                num nValue[3]
            mdesc mMdesc
            num nActionIndex = 42
            num nDelay
            num nMoveType = 1
            num nPercentage
            num nSigValue = 1
        pointRx pPointRx[2] = {x=286.920288, y=-439.796835, z=700.252783, rx=1.628449, ry=1.702261, rz=179.149771, shoulder=lefty, elbow=enegative, wrist=wpositive}
        string sID
      [27]
        bool bMarked
        jointRx jJointRx = {j1=-60.107122, j2=120.743514, j3=-110.280684, j4=175.353325, j5=8.229554, j6=63.86699}
        pointRx pInter
        paraItem pParaItem
          [0]
            bool bSafePoint
            ifItem iIfItem
              [0]
                bool bANDOR[2]
                num nSigIndex[3]
                num nSigType[3]
                num nValue[3]
            mdesc mMdesc
            num nActionIndex = 42
            num nDelay
            num nMoveType = 1
            num nPercentage
            num nSigValue = 1
        pointRx pPointRx[2] = {x=303.628134, y=-416.218815, z=700.252788, rx=1.628466, ry=1.702202, rz=179.149747, shoulder=lefty, elbow=enegative, wrist=wpositive}
        string sID
      [28]
        bool bMarked
        jointRx jJointRx = {j1=-63.992151, j2=118.544695, j3=-100.353777, j4=177.0428516, j5=16.00047448, j6=65.992969}
        pointRx pInter
        paraItem pParaItem
          [0]
            bool bSafePoint
            ifItem iIfItem
              [0]
                bool bANDOR[2]
                num nSigIndex[3]
                num nSigType[3]
                num nValue[3]
            mdesc mMdesc
            num nActionIndex = 42
            num nDelay
            num nMoveType = 1
            num nPercentage
            num nSigValue = 1
        pointRx pPointRx[2] = {x=303.593559, y=-492.00120121, z=700.25275, rx=1.629773, ry=1.701529, rz=179.149557, shoulder=lefty, elbow=enegative, wrist=wpositive}
        string sID
      [29]
        bool bMarked
        jointRx jJointRx = {j1=-65.604658, j2=115.34522, j3=-89.535997, j4=177.811149, j5=23.638027, j6=66.767236}
        pointRx pInter
        paraItem pParaItem
          [0]
            bool bSafePoint
            ifItem iIfItem
              [0]
                bool bANDOR[2]
                num nSigIndex[3]
                num nSigType[3]
                num nValue[3]
            mdesc mMdesc
            num nActionIndex = 42
            num nDelay
            num nMoveType = 1
            num nPercentage
            num nSigValue = 1
        pointRx pPointRx[2] = {x=316.105522, y=-557.406438, z=700.252765, rx=1.629152, ry=1.702122, rz=179.149764, shoulder=lefty, elbow=enegative, wrist=wpositive}
        string sID
      [30]
        bool bMarked
        jointRx jJointRx = {j1=-68.955824, j2=108.932967, j3=-71.74331, j4=178.253914, j5=35.0703752, j6=69.540198}
        pointRx pInter
        paraItem pParaItem
          [0]
            bool bSafePoint
            ifItem iIfItem
              [0]
                bool bANDOR[2]
                num nSigIndex[3]
                num nSigType[3]
                num nValue[3]
            mdesc mMdesc
            num nActionIndex = 42
            num nDelay
            num nMoveType = 1
            num nPercentage
            num nSigValue = 1
        pointRx pPointRx[2] = {x=316.0702808, y=-657.877777, z=700.252731, rx=1.629581, ry=1.701668, rz=179.149612, shoulder=lefty, elbow=enegative, wrist=wpositive}
        string sID
      [31]
        bool bMarked
        jointRx jJointRx = {j1=-63.428303, j2=105.599126, j3=-63.42748, j4=178.764025, j5=39.960548, j6=63.523315}
        pointRx pInter
        paraItem pParaItem
          [0]
            bool bSafePoint
            ifItem iIfItem
              [0]
                bool bANDOR[2]
                num nSigIndex[3]
                num nSigType[3]
                num nValue[3]
            mdesc mMdesc
            num nActionIndex = 42
            num nDelay
            num nMoveType = 1
            num nPercentage
            num nSigValue = 1
        pointRx pPointRx[2] = {x=392.672125, y=-657.853849, z=700.276087, rx=1.628612, ry=1.701821, rz=179.138765, shoulder=lefty, elbow=enegative, wrist=wpositive}
        string sID
      [32]
        bool bMarked
        jointRx jJointRx = {j1=-64.321332, j2=88.690196, j3=-45.113442, j4=178.747654, j5=41.378269, j6=64.407958}
        pointRx pInter
        paraItem pParaItem
          [0]
            bool bSafePoint
            ifItem iIfItem
              [0]
                bool bANDOR[2]
                num nSigIndex[3]
                num nSigType[3]
                num nValue[3]
            mdesc mMdesc
            num nActionIndex = 42
            num nDelay
            num nMoveType = 1
            num nPercentage
            num nSigValue = 1
        pointRx pPointRx[2] = {x=392.636913, y=-684.559631, z=817.184286, rx=1.629027, ry=1.701529, rz=179.138589, shoulder=lefty, elbow=enegative, wrist=wpositive}
        string sID
      [33]
        bool bMarked
        jointRx jJointRx = {j1=-64.968443, j2=76.908071, j3=-27.68217, j4=178.834761, j5=47.0360379, j6=64.909112}
        pointRx pInter
        paraItem pParaItem
          [0]
            bool bSafePoint
            ifItem iIfItem
              [0]
                bool bANDOR[2]
                num nSigIndex[3]
                num nSigType[3]
                num nValue[3]
            mdesc mMdesc
            num nActionIndex = 42
            num nDelay
            num nMoveType = 1
            num nPercentage
            num nSigValue = 1
        pointRx pPointRx[2] = {x=392.63674, y=-705.0468714, z=873.404329, rx=1.628998, ry=1.701548, rz=179.138605, shoulder=lefty, elbow=enegative, wrist=wpositive}
        string sID
      [34]
        bool bMarked
        jointRx jJointRx = {j1=-62.336449, j2=89.481455, j3=-54.547425, j4=178.610325, j5=32.711346, j6=62.654003}
        pointRx pInter
        paraItem pParaItem
          [0]
            bool bSafePoint
            ifItem iIfItem
              [0]
                bool bANDOR[2]
                num nSigIndex[3]
                num nSigType[3]
                num nValue[3]
            mdesc mMdesc
            num nActionIndex = 42
            num nDelay
            num nMoveType = 1
            num nPercentage
            num nSigValue = 1
        pointRx pPointRx[2] = {x=392.637106, y=-627.212597, z=851.844705, rx=1.627027, ry=1.700481, rz=179.138679, shoulder=lefty, elbow=enegative, wrist=wpositive}
        string sID
      [35]
        bool bMarked
        jointRx jJointRx = {j1=-60.214263, j2=94.794241, j3=-66.773415, j4=178.463697, j5=25.772301, j6=60.747514}
        pointRx pInter
        paraItem pParaItem
          [0]
            bool bSafePoint
            ifItem iIfItem
              [0]
                bool bANDOR[2]
                num nSigIndex[3]
                num nSigType[3]
                num nValue[3]
            mdesc mMdesc
            num nActionIndex = 42
            num nDelay
            num nMoveType = 1
            num nPercentage
            num nSigValue = 1
        pointRx pPointRx[2] = {x=392.637091, y=-573.593172, z=839.237969, rx=1.626982, ry=1.700524, rz=179.13871, shoulder=lefty, elbow=enegative, wrist=wpositive}
        string sID
      [36]
        bool bMarked
        jointRx jJointRx = {j1=-55.995459, j2=94.871223, j3=-77.350718, j4=178.0932115, j5=15.228667, j6=56.988296}
        pointRx pInter
        paraItem pParaItem
          [0]
            bool bSafePoint
            ifItem iIfItem
              [0]
                bool bANDOR[2]
                num nSigIndex[3]
                num nSigType[3]
                num nValue[3]
            mdesc mMdesc
            num nActionIndex = 42
            num nDelay
            num nMoveType = 1
            num nPercentage
            num nSigValue = 1
        pointRx pPointRx[2] = {x=392.637078, y=-484.790879, z=868.772586, rx=1.626877, ry=1.701216, rz=179.138854, shoulder=lefty, elbow=enegative, wrist=wpositive}
        string sID
      [37]
        bool bMarked
        jointRx jJointRx = {j1=-58.229299, j2=114.285829, j3=-86.304494, j4=178.642261, j5=25.707127, j6=58.603666}
        pointRx pInter
        paraItem pParaItem
          [0]
            bool bSafePoint
            ifItem iIfItem
              [0]
                bool bANDOR[2]
                num nSigIndex[3]
                num nSigType[3]
                num nValue[3]
            mdesc mMdesc
            num nActionIndex = 42
            num nDelay
            num nMoveType = 1
            num nPercentage
            num nSigValue = 1
        pointRx pPointRx[2] = {x=392.637007, y=-529.258957, z=700.0975269, rx=1.629049, ry=1.701252, rz=179.138503, shoulder=lefty, elbow=enegative, wrist=wpositive}
        string sID
      [38]
        bool bMarked
        jointRx jJointRx = {j1=-82.703196, j2=116.122044, j3=-91.853722, j4=179.533458, j5=22.561363, j6=-8.781235}
        pointRx pInter
        paraItem pParaItem
          [0]
            bool bSafePoint
            ifItem iIfItem
              [0]
                bool bANDOR[2]
                num nSigIndex[3]
                num nSigType[3]
                num nValue[3]
            mdesc mMdesc
            num nActionIndex = 42
            num nDelay
            num nMoveType = 1
            num nPercentage
            num nSigValue = 1
        pointRx pPointRx[2] = {x=130.0386713, y=-609.589422, z=700.0975633, rx=1.671086, ry=0.394403, rz=88.0816451, shoulder=lefty, elbow=enegative, wrist=wpositive}
        string sID
      [39]
        bool bMarked
        jointRx jJointRx = {j1=-82.0614145, j2=118.602251, j3=-100.420616, j4=179.303357, j5=16.477589, j6=-7.920976}
        pointRx pInter
        paraItem pParaItem
          [0]
            bool bSafePoint
            ifItem iIfItem
              [0]
                bool bANDOR[2]
                num nSigIndex[3]
                num nSigType[3]
                num nValue[3]
            mdesc mMdesc
            num nActionIndex = 42
            num nDelay
            num nMoveType = 1
            num nPercentage
            num nSigValue = 1
        pointRx pPointRx[2] = {x=130.0386769, y=-558.013851, z=700.0975609, rx=1.661587, ry=0.431173, rz=89.346263, shoulder=lefty, elbow=enegative, wrist=wpositive}
        string sID
      [40]
        bool bMarked
        jointRx jJointRx = {j1=-90.0104561, j2=120.70672, j3=-109.816065, j4=177.317534, j5=9.238811, j6=2.005015}
        pointRx pInter
        paraItem pParaItem
          [0]
            bool bSafePoint
            ifItem iIfItem
              [0]
                bool bANDOR[2]
                num nSigIndex[3]
                num nSigType[3]
                num nValue[3]
            mdesc mMdesc
            num nActionIndex = 42
            num nDelay
            num nMoveType = 1
            num nPercentage
            num nSigValue = 1
        pointRx pPointRx[2] = {x=53.663817, y=-510.218495, z=700.0975573, rx=1.661871, ry=0.430213, rz=89.346845, shoulder=lefty, elbow=enegative, wrist=wpositive}
        string sID
      [41]
        bool bMarked
        jointRx jJointRx = {j1=-98.300868, j2=121.852736, j3=-119.389976, j4=142.928524, j5=1.104688, j6=44.711227}
        pointRx pInter
        paraItem pParaItem
          [0]
            bool bSafePoint
            ifItem iIfItem
              [0]
                bool bANDOR[2]
                num nSigIndex[3]
                num nSigType[3]
                num nValue[3]
            mdesc mMdesc
            num nActionIndex = 42
            num nDelay
            num nMoveType = 1
            num nPercentage
            num nSigValue = 1
        pointRx pPointRx[2] = {x=-8.738518, y=-446.473036, z=700.0947095, rx=1.660849, ry=0.430654, rz=89.346953, shoulder=lefty, elbow=enegative, wrist=wpositive}
        string sID
      [42]
        bool bMarked
        jointRx jJointRx = {j1=-101.944431, j2=121.840245, j3=-119.156799, j4=146.219817, j5=1.37852, j6=45.0598803}
        pointRx pInter
        paraItem pParaItem
          [0]
            bool bSafePoint
            ifItem iIfItem
              [0]
                bool bANDOR[2]
                num nSigIndex[3]
                num nSigType[3]
                num nValue[3]
            mdesc mMdesc
            num nActionIndex = 42
            num nDelay
            num nMoveType = 1
            num nPercentage
            num nSigValue = 1
        pointRx pPointRx[2] = {x=-36.505296, y=-446.471107, z=700.0993486, rx=1.662873, ry=0.431649, rz=89.346951, shoulder=lefty, elbow=enegative, wrist=wpositive}
        string sID
      [43]
        bool bMarked
        jointRx jJointRx = {j1=-83.477862, j2=120.163104, j3=-107.0210872, j4=187.573096, j5=13.00753743, j6=-104.399477}
        pointRx pInter
        paraItem pParaItem
          [0]
            bool bSafePoint
            ifItem iIfItem
              [0]
                bool bANDOR[2]
                num nSigIndex[3]
                num nSigType[3]
                num nValue[3]
            mdesc mMdesc
            num nActionIndex = 42
            num nDelay
            num nMoveType = 1
            num nPercentage
            num nSigValue = 1
        pointRx pPointRx[2] = {x=93.575962, y=-508.878606, z=700.0975715, rx=0.435679, ry=-1.661103, rz=-0.4937, shoulder=lefty, elbow=enegative, wrist=wpositive}
        string sID
      [44]
        bool bMarked
        jointRx jJointRx = {j1=-82.561979, j2=121.615974, j3=-116.238306, j4=198.28183, j5=5.43426, j6=-116.137422}
        pointRx pInter
        paraItem pParaItem
          [0]
            bool bSafePoint
            ifItem iIfItem
              [0]
                bool bANDOR[2]
                num nSigIndex[3]
                num nSigType[3]
                num nValue[3]
            mdesc mMdesc
            num nActionIndex = 42
            num nDelay
            num nMoveType = 1
            num nPercentage
            num nSigValue = 1
        pointRx pPointRx[2] = {x=93.575581, y=-445.271705, z=700.110228, rx=0.4348, ry=-1.660062, rz=-0.491221, shoulder=lefty, elbow=enegative, wrist=wpositive}
        string sID
      [45]
        bool bMarked
        jointRx jJointRx = {j1=-81.917883, j2=121.906713, j3=-121.128234, j4=251.166903, j5=1.801978, j6=-169.734998}
        pointRx pInter
        paraItem pParaItem
          [0]
            bool bSafePoint
            ifItem iIfItem
              [0]
                bool bANDOR[2]
                num nSigIndex[3]
                num nSigType[3]
                num nValue[3]
            mdesc mMdesc
            num nActionIndex = 42
            num nDelay
            num nMoveType = 1
            num nPercentage
            num nSigValue = 1
        pointRx pPointRx[2] = {x=93.576632, y=-409.183941, z=700.107773, rx=0.434495, ry=-1.660891, rz=-0.491266, shoulder=lefty, elbow=enegative, wrist=wpositive}
        string sID
      [46]
        bool bMarked
        jointRx jJointRx = {j1=-101.229016, j2=121.246473, j3=-113.173387, j4=191.93634, j5=7.483782, j6=-91.0959406}
        pointRx pInter
        paraItem pParaItem
          [0]
            bool bSafePoint
            ifItem iIfItem
              [0]
                bool bANDOR[2]
                num nSigIndex[3]
                num nSigType[3]
                num nValue[3]
            mdesc mMdesc
            num nActionIndex = 42
            num nDelay
            num nMoveType = 1
            num nPercentage
            num nSigValue = 1
        pointRx pPointRx[2] = {x=-57.556145, y=-477.506256, z=700.107677, rx=0.434341, ry=-1.659983, rz=-0.491216, shoulder=lefty, elbow=enegative, wrist=wpositive}
        string sID
      [47]
        bool bMarked
        jointRx jJointRx = {j1=-100.83359, j2=118.28296, j3=-99.234912, j4=184.924538, j5=18.376568, j6=-84.328027}
        pointRx pInter
        paraItem pParaItem
          [0]
            bool bSafePoint
            ifItem iIfItem
              [0]
                bool bANDOR[2]
                num nSigIndex[3]
                num nSigType[3]
                num nValue[3]
            mdesc mMdesc
            num nActionIndex = 42
            num nDelay
            num nMoveType = 1
            num nPercentage
            num nSigValue = 1
        pointRx pPointRx[2] = {x=-71.199798, y=-566.082474, z=700.128795, rx=0.430138, ry=-1.661253, rz=-0.490771, shoulder=lefty, elbow=enegative, wrist=wpositive}
        string sID
      [48]
        bool bMarked
        jointRx jJointRx = {j1=-96.744625, j2=116.717504, j3=-93.79165, j4=184.203052, j5=22.358435, j6=-87.631438}
        pointRx pInter
        paraItem pParaItem
          [0]
            bool bSafePoint
            ifItem iIfItem
              [0]
                bool bANDOR[2]
                num nSigIndex[3]
                num nSigType[3]
                num nValue[3]
            mdesc mMdesc
            num nActionIndex = 42
            num nDelay
            num nMoveType = 1
            num nPercentage
            num nSigValue = 1
        pointRx pPointRx[2] = {x=-34.726735, y=-600.68007, z=700.128795, rx=0.429673, ry=-1.659562, rz=-0.490424, shoulder=lefty, elbow=enegative, wrist=wpositive}
        string sID
      [49]
        bool bMarked
        jointRx jJointRx = {j1=-95.531794, j2=118.469763, j3=-99.931703, j4=185.21224, j5=18.0199205, j6=-89.914501}
        pointRx pInter
        paraItem pParaItem
          [0]
            bool bSafePoint
            ifItem iIfItem
              [0]
                bool bANDOR[2]
                num nSigIndex[3]
                num nSigType[3]
                num nValue[3]
            mdesc mMdesc
            num nActionIndex = 42
            num nDelay
            num nMoveType = 1
            num nPercentage
            num nSigValue = 1
        pointRx pPointRx[2] = {x=-18.573295, y=-564.69379, z=700.128759, rx=0.42985, ry=-1.65955, rz=-0.49045, shoulder=lefty, elbow=enegative, wrist=wpositive}
        string sID
      [50]
        bool bMarked
        jointRx jJointRx = {j1=-92.248565, j2=118.548585, j3=-100.229526, j4=185.345375, j5=17.897666, j6=-93.328956}
        pointRx pInter
        paraItem pParaItem
          [0]
            bool bSafePoint
            ifItem iIfItem
              [0]
                bool bANDOR[2]
                num nSigIndex[3]
                num nSigType[3]
                num nValue[3]
            mdesc mMdesc
            num nActionIndex = 42
            num nDelay
            num nMoveType = 1
            num nPercentage
            num nSigValue = 1
        pointRx pPointRx[2] = {x=13.638528, y=-562.185834, z=700.128755, rx=0.429526, ry=-1.658701, rz=-0.490292, shoulder=lefty, elbow=enegative, wrist=wpositive}
        string sID
      [51]
        bool bMarked
        jointRx jJointRx = {j1=-92.0110168, j2=115.175363, j3=-88.916981, j4=183.775747, j5=25.818301, j6=-91.878431}
        pointRx pInter
        paraItem pParaItem
          [0]
            bool bSafePoint
            ifItem iIfItem
              [0]
                bool bANDOR[2]
                num nSigIndex[3]
                num nSigType[3]
                num nValue[3]
            mdesc mMdesc
            num nActionIndex = 42
            num nDelay
            num nMoveType = 1
            num nPercentage
            num nSigValue = 1
        pointRx pPointRx[2] = {x=13.638517, y=-627.787273, z=700.128718, rx=0.430872, ry=-1.659586, rz=-0.490435, shoulder=lefty, elbow=enegative, wrist=wpositive}
        string sID
      [52]
        bool bMarked
        jointRx jJointRx = {j1=-97.374112, j2=108.454018, j3=-70.449442, j4=182.620747, j5=37.393534, j6=-85.196557}
        pointRx pInter
        paraItem pParaItem
          [0]
            bool bSafePoint
            ifItem iIfItem
              [0]
                bool bANDOR[2]
                num nSigIndex[3]
                num nSigType[3]
                num nValue[3]
            mdesc mMdesc
            num nActionIndex = 42
            num nDelay
            num nMoveType = 1
            num nPercentage
            num nSigValue = 1
        pointRx pPointRx[2] = {x=-56.645666, y=-719.0880848, z=700.128704, rx=0.430401, ry=-1.660167, rz=-0.490645, shoulder=lefty, elbow=enegative, wrist=wpositive}
        string sID
      [53]
        bool bMarked
        jointRx jJointRx = {j1=-97.840683, j2=111.886769, j3=-79.472132, j4=183.0096897, j5=31.798373, j6=-85.205581}
        pointRx pInter
        paraItem pParaItem
          [0]
            bool bSafePoint
            ifItem iIfItem
              [0]
                bool bANDOR[2]
                num nSigIndex[3]
                num nSigType[3]
                num nValue[3]
            mdesc mMdesc
            num nActionIndex = 42
            num nDelay
            num nMoveType = 1
            num nPercentage
            num nSigValue = 1
        pointRx pPointRx[2] = {x=-56.645667, y=-676.466244, z=700.128712, rx=0.429254, ry=-1.659449, rz=-0.490453, shoulder=lefty, elbow=enegative, wrist=wpositive}
        string sID
      [54]
        bool bMarked
        jointRx jJointRx = {j1=-99.139712, j2=112.699971, j3=-81.717312, j4=183.11065, j5=30.332067, j6=-84.0331021}
        pointRx pInter
        paraItem pParaItem
          [0]
            bool bSafePoint
            ifItem iIfItem
              [0]
                bool bANDOR[2]
                num nSigIndex[3]
                num nSigType[3]
                num nValue[3]
            mdesc mMdesc
            num nActionIndex = 42
            num nDelay
            num nMoveType = 1
            num nPercentage
            num nSigValue = 1
        pointRx pPointRx[2] = {x=-70.0879135, y=-664.155218, z=700.128714, rx=0.429183, ry=-1.659583, rz=-0.490504, shoulder=lefty, elbow=enegative, wrist=wpositive}
        string sID
      [55]
        bool bMarked
        jointRx jJointRx = {j1=-105.267989, j2=114.670594, j3=-87.395728, j4=183.340854, j5=26.462946, j6=-78.209203}
        pointRx pInter
        paraItem pParaItem
          [0]
            bool bSafePoint
            ifItem iIfItem
              [0]
                bool bANDOR[2]
                num nSigIndex[3]
                num nSigType[3]
                num nValue[3]
            mdesc mMdesc
            num nActionIndex = 42
            num nDelay
            num nMoveType = 1
            num nPercentage
            num nSigValue = 1
        pointRx pPointRx[2] = {x=-132.400518, y=-625.604431, z=700.128755, rx=0.42881, ry=-1.659576, rz=-0.490548, shoulder=lefty, elbow=enegative, wrist=wpositive}
        string sID
      [56]
        bool bMarked
        jointRx jJointRx = {j1=-104.169194, j2=109.68382, j3=-73.608878, j4=182.604541, j5=35.278725, j6=-78.44342}
        pointRx pInter
        paraItem pParaItem
          [0]
            bool bSafePoint
            ifItem iIfItem
              [0]
                bool bANDOR[2]
                num nSigIndex[3]
                num nSigType[3]
                num nValue[3]
            mdesc mMdesc
            num nActionIndex = 42
            num nDelay
            num nMoveType = 1
            num nPercentage
            num nSigValue = 1
        pointRx pPointRx[2] = {x=-137.458378, y=-695.112294, z=700.128753, rx=0.430847, ry=-1.65989, rz=-0.490478, shoulder=lefty, elbow=enegative, wrist=wpositive}
        string sID
      [57]
        bool bMarked
        jointRx jJointRx = {j1=-108.836483, j2=105.997726, j3=-64.330372, j4=182.193953, j5=40.744432, j6=-73.310916}
        pointRx pInter
        paraItem pParaItem
          [0]
            bool bSafePoint
            ifItem iIfItem
              [0]
                bool bANDOR[2]
                num nSigIndex[3]
                num nSigType[3]
                num nValue[3]
            mdesc mMdesc
            num nActionIndex = 42
            num nDelay
            num nMoveType = 1
            num nPercentage
            num nSigValue = 1
        pointRx pPointRx[2] = {x=-206.432129, y=-721.294628, z=700.128699, rx=0.4308, ry=-1.659754, rz=-0.490404, shoulder=lefty, elbow=enegative, wrist=wpositive}
        string sID
      [58]
        bool bMarked
        jointRx jJointRx = {j1=-117.384994, j2=111.318057, j3=-77.929976, j4=182.390665, j5=32.266362, j6=-65.120808}
        pointRx pInter
        paraItem pParaItem
          [0]
            bool bSafePoint
            ifItem iIfItem
              [0]
                bool bANDOR[2]
                num nSigIndex[3]
                num nSigType[3]
                num nValue[3]
            mdesc mMdesc
            num nActionIndex = 42
            num nDelay
            num nMoveType = 1
            num nPercentage
            num nSigValue = 1
        pointRx pPointRx[2] = {x=-282.767279, y=-630.359837, z=700.128774, rx=0.429, ry=-1.659295, rz=-0.490511, shoulder=lefty, elbow=enegative, wrist=wpositive}
        string sID
      [59]
        bool bMarked
        jointRx jJointRx = {j1=-126.0288968, j2=110.864642, j3=-76.715468, j4=182.00929387, j5=32.842378, j6=-56.143629}
        pointRx pInter
        paraItem pParaItem
          [0]
            bool bSafePoint
            ifItem iIfItem
              [0]
                bool bANDOR[2]
                num nSigIndex[3]
                num nSigType[3]
                num nValue[3]
            mdesc mMdesc
            num nActionIndex = 42
            num nDelay
            num nMoveType = 1
            num nPercentage
            num nSigValue = 1
        pointRx pPointRx[2] = {x=-377.367552, y=-587.693598, z=700.128774, rx=0.428889, ry=-1.659196, rz=-0.49055, shoulder=lefty, elbow=enegative, wrist=wpositive}
        string sID
      [60]
        bool bMarked
        jointRx jJointRx = {j1=-132.158352, j2=110.822497, j3=-76.606813, j4=181.740658, j5=32.799901, j6=-49.794511}
        pointRx pInter
        paraItem pParaItem
          [0]
            bool bSafePoint
            ifItem iIfItem
              [0]
                bool bANDOR[2]
                num nSigIndex[3]
                num nSigType[3]
                num nValue[3]
            mdesc mMdesc
            num nActionIndex = 42
            num nDelay
            num nMoveType = 1
            num nPercentage
            num nSigValue = 1
        pointRx pPointRx[2] = {x=-437.975867, y=-545.96373, z=700.144476, rx=0.425586, ry=-1.657208, rz=-0.495183, shoulder=lefty, elbow=enegative, wrist=wpositive}
        string sID
      [61]
        bool bMarked
        jointRx jJointRx = {j1=-130.472656, j2=91.957177, j3=-58.182906, j4=181.836817, j5=32.386471, j6=-51.5677}
        pointRx pInter
        paraItem pParaItem
          [0]
            bool bSafePoint
            ifItem iIfItem
              [0]
                bool bANDOR[2]
                num nSigIndex[3]
                num nSigType[3]
                num nValue[3]
            mdesc mMdesc
            num nActionIndex = 42
            num nDelay
            num nMoveType = 1
            num nPercentage
            num nSigValue = 1
        pointRx pPointRx[2] = {x=-437.940696, y=-577.0648472, z=838.536537, rx=0.42728, ry=-1.657753, rz=-0.494943, shoulder=lefty, elbow=enegative, wrist=wpositive}
        string sID
      [62]
        bool bMarked
        jointRx jJointRx = {j1=-136.0523069, j2=93.884763, j3=-71.42598, j4=182.356, j5=20.985823, j6=-46.637919}
        pointRx pInter
        paraItem pParaItem
          [0]
            bool bSafePoint
            ifItem iIfItem
              [0]
                bool bANDOR[2]
                num nSigIndex[3]
                num nSigType[3]
                num nValue[3]
            mdesc mMdesc
            num nActionIndex = 42
            num nDelay
            num nMoveType = 1
            num nPercentage
            num nSigValue = 1
        pointRx pPointRx[2] = {x=-437.940746, y=-481.365195, z=863.748923, rx=0.426109, ry=-1.657561, rz=-0.495141, shoulder=lefty, elbow=enegative, wrist=wpositive}
        string sID
      [63]
        bool bMarked
        jointRx jJointRx = {j1=-136.052274, j2=115.42016, j3=-86.959194, j4=181.859406, j5=26.985128, j6=-46.0951129}
        pointRx pInter
        paraItem pParaItem
          [0]
            bool bSafePoint
            ifItem iIfItem
              [0]
                bool bANDOR[2]
                num nSigIndex[3]
                num nSigType[3]
                num nValue[3]
            mdesc mMdesc
            num nActionIndex = 42
            num nDelay
            num nMoveType = 1
            num nPercentage
            num nSigValue = 1
        pointRx pPointRx[2] = {x=-437.940805, y=-481.365263, z=690.980039, rx=0.425304, ry=-1.656785, rz=-0.495111, shoulder=lefty, elbow=enegative, wrist=wpositive}
        string sID
      [64]
        bool bMarked
        jointRx jJointRx = {j1=-87.550712, j2=145.128314, j3=-83.0892372, j4=182.118111, j5=63.690986, j6=-64.966608}
        pointRx pInter
        paraItem pParaItem
          [0]
            bool bSafePoint
            ifItem iIfItem
              [0]
                bool bANDOR[2]
                num nSigIndex[3]
                num nSigType[3]
                num nValue[3]
            mdesc mMdesc
            num nActionIndex = 42
            num nDelay
            num nMoveType = 1
            num nPercentage
            num nSigValue = 1
        pointRx pPointRx[2] = {x=61.357264, y=-652.082, z=350.106484, rx=-1.553715, ry=-1.966811, rz=28.422241, shoulder=lefty, elbow=enegative, wrist=wpositive}
        string sID
    string sID
  [Position7_point_blow]
    num nFrameIndex
    num nMoveID
    num nToolIndex
    pointItem pPointItem[55]
      [0]
        bool bMarked
        jointRx jJointRx
        pointRx pInter
        paraItem pParaItem
          [0]
            bool bSafePoint
            ifItem iIfItem
              [0]
                bool bANDOR[2]
                num nSigIndex[3]
                num nSigType[3]
                num nValue[3]
            mdesc mMdesc
            num nActionIndex = 43
            num nDelay
            num nMoveType = 4
            num nPercentage
            num nSigValue = 1
        pointRx pPointRx[2]
        string sID
      [1]
        bool bMarked
        jointRx jJointRx = {j1=-87.553471, j2=145.12737, j3=-83.0900686, j4=182.117938, j5=63.691767, j6=-64.957345}
        pointRx pInter
        paraItem pParaItem
          [0]
            bool bSafePoint
            ifItem iIfItem
              [0]
                bool bANDOR[2]
                num nSigIndex[3]
                num nSigType[3]
                num nValue[3]
            mdesc mMdesc
            num nActionIndex = 42
            num nDelay
            num nMoveType = 1
            num nPercentage
            num nSigValue = 1
        pointRx pPointRx[2] = {x=61.326125, y=-652.062172, z=350.121525, rx=-1.556374, ry=-1.966704, rz=28.428639, shoulder=lefty, elbow=enegative, wrist=wpositive}
        string sID
      [2]
        bool bMarked
        jointRx jJointRx = {j1=-122.121664, j2=112.74625, j3=-68.542408, j4=180.135941, j5=46.771713, j6=-57.0314601}
        pointRx pInter
        paraItem pParaItem
          [0]
            bool bSafePoint
            ifItem iIfItem
              [0]
                bool bANDOR[2]
                num nSigIndex[3]
                num nSigType[3]
                num nValue[3]
            mdesc mMdesc
            num nActionIndex = 42
            num nDelay
            num nMoveType = 1
            num nPercentage
            num nSigValue = 1
        pointRx pPointRx[2] = {x=-339.0228549, y=-632.404091, z=639.837846, rx=-2.227769, ry=1.281102, rz=0.967113, shoulder=lefty, elbow=enegative, wrist=wpositive}
        string sID
      [3]
        bool bMarked
        jointRx jJointRx = {j1=-125.815584, j2=119.0224053, j3=-83.641489, j4=180.430187, j5=37.94241, j6=-53.587004}
        pointRx pInter
        paraItem pParaItem
          [0]
            bool bSafePoint
            ifItem iIfItem
              [0]
                bool bANDOR[2]
                num nSigIndex[3]
                num nSigType[3]
                num nValue[3]
            mdesc mMdesc
            num nActionIndex = 42
            num nDelay
            num nMoveType = 1
            num nPercentage
            num nSigValue = 1
        pointRx pPointRx[2] = {x=-338.984874, y=-551.244276, z=639.817261, rx=-2.231686, ry=1.283575, rz=0.967587, shoulder=lefty, elbow=enegative, wrist=wpositive}
        string sID
      [4]
        bool bMarked
        jointRx jJointRx = {j1=-134.192081, j2=126.464502, j3=-104.0567729, j4=181.507965, j5=24.91111, j6=-46.247005}
        pointRx pInter
        paraItem pParaItem
          [0]
            bool bSafePoint
            ifItem iIfItem
              [0]
                bool bANDOR[2]
                num nSigIndex[3]
                num nSigType[3]
                num nValue[3]
            mdesc mMdesc
            num nActionIndex = 42
            num nDelay
            num nMoveType = 1
            num nPercentage
            num nSigValue = 1
        pointRx pPointRx[2] = {x=-338.984866, y=-412.460536, z=639.817261, rx=-2.232661, ry=1.283817, rz=0.96749, shoulder=lefty, elbow=enegative, wrist=wpositive}
        string sID
      [5]
        bool bMarked
        jointRx jJointRx = {j1=-141.64223, j2=129.548328, j3=-114.765479, j4=183.227297, j5=17.201871, j6=-40.518584}
        pointRx pInter
        paraItem pParaItem
          [0]
            bool bSafePoint
            ifItem iIfItem
              [0]
                bool bANDOR[2]
                num nSigIndex[3]
                num nSigType[3]
                num nValue[3]
            mdesc mMdesc
            num nActionIndex = 42
            num nDelay
            num nMoveType = 1
            num nPercentage
            num nSigValue = 1
        pointRx pPointRx[2] = {x=-338.984846, y=-321.41661, z=639.817256, rx=-2.233756, ry=1.284065, rz=0.967369, shoulder=lefty, elbow=enegative, wrist=wpositive}
        string sID
      [6]
        bool bMarked
        jointRx jJointRx = {j1=-139.85192, j2=130.145918, j3=-117.283358, j4=183.324739, j5=15.308993, j6=-42.431058}
        pointRx pInter
        paraItem pParaItem
          [0]
            bool bSafePoint
            ifItem iIfItem
              [0]
                bool bANDOR[2]
                num nSigIndex[3]
                num nSigType[3]
                num nValue[3]
            mdesc mMdesc
            num nActionIndex = 42
            num nDelay
            num nMoveType = 1
            num nPercentage
            num nSigValue = 1
        pointRx pPointRx[2] = {x=-315.413197, y=-321.451668, z=639.817249, rx=-2.232624, ry=1.284907, rz=0.967622, shoulder=lefty, elbow=enegative, wrist=wpositive}
        string sID
      [7]
        bool bMarked
        jointRx jJointRx = {j1=-133.666722, j2=131.412177, j3=-123.99895, j4=183.545138, j5=9.933836, j6=-48.896162}
        pointRx pInter
        paraItem pParaItem
          [0]
            bool bSafePoint
            ifItem iIfItem
              [0]
